Fanuc KAREL source: KT00606.KL

PROGRAM KT00606
%NOLOCKGROUP
VAR
  I1: INTEGER
  I2: INTEGER
  OUT: BOOLEAN
BEGIN
  I1 = 2
  I2 = 3
  I1 = 2
  I2 = 3
  OUT = - I1
END KT00606
